Fanuc KAREL source: KB00075.KL

PROGRAM KB00075
%NOLOCKGROUP
%ENVIRONMENT FDEV
VAR
  P1: STRING[80]
  P2: STRING[80]
  P3: BOOLEAN
  P4: INTEGER
BEGIN
  P1 = 'A'
  P2 = 'A'
  P3 = TRUE
  P4 = 1
  FORMAT_DEV(P1, P2, P3, P4)
END KB00075
